(* IEC 61131-3 sources: plcassist-cli/packages/volt-lsp-iec/test-corpus/awa-palletizer/Device/Plc Logic/Application/Library Manager/(unresolved)/sysprocess interfaces, 1 file *)

(* ---- GLOBAL_CONSTANTS.gvl ---- *)
VAR_GLOBAL
	SYSPROCESS_INVALID_HANDLE : UDINT := 16#FFFFFFFF;
	SYSPROCESS_CREATEFLAG_HIDDEN : UDINT := 16#1;
	SYSPROCESS_CREATEFLAG_INTERACTIVE : UDINT := 16#2;
	SYSPROCESS_CREATEFLAG_CREATESUSPENDED : UDINT := 16#4;
END_VAR
